(* IEC 61131-3 sources: Elmo_Master/Lasal_PRG/Welcon8Axis_EtherCAT_Test_With_RobotAxis/Class/HwControl (part 3) *)

      // safety settings
      //*********************************************************************************************
      HWC_PARA_IDX_SAFETY:

        // SubIndex
        //----------------------------------------------------------------------------------
        case SubIndex of

          //--------------------------------------------------------------------------------
          HWC_PARA_SUBIDX_SAFETY_UDP_TIME: // override cycle interval for UDP communication

            SafetyManager.GetUdpParameters(pCycleTime:=pValue$^UDINT, pTimeout:=NIL);

            Retcode := 0; // success

          //--------------------------------------------------------------------------------
          HWC_PARA_SUBIDX_SAFETY_UDP_TIMEOUT: // override timeout value for UDP communication

            SafetyManager.GetUdpParameters(pCycleTime:=NIL, pTimeout:=pValue$^UDINT);

            Retcode := 0; // success

          //--------------------------------------------------------------------------------
          else
            Retcode := -2;  // invalid SubIdx
          end_case;
    //--------------------------------------------------------------------------------
    else
      Retcode := -1;  // invalid Index
    end_case;
  end_if;

END_FUNCTION

FUNCTION GLOBAL HwControl::SetPara
	VAR_INPUT
		Index 	: DINT;
		SubIndex 	: DINT;
		Value 	: DINT;
	END_VAR
	VAR_OUTPUT
		Retcode 	: DINT;
	END_VAR

  // init returncode with invalid index
  Retcode := -1;

  // Index
  //***********************************************************************************************
  case Index of

    // safety settings
    //*********************************************************************************************
    HWC_PARA_IDX_SAFETY:

      // SubIndex
      //----------------------------------------------------------------------------------
      case SubIndex of

        //--------------------------------------------------------------------------------
        HWC_PARA_SUBIDX_SAFETY_UDP_TIME: // override cycle interval for UDP communication

          // value needs to be at least 2ms
          if Value >= 2 then
            // check if the init phase hasn't been finished yet
            if (us_InitCounter < 12) then
              SafetyManager.SetUdpParameters(pCycleTime:=(#Value)$^UDINT, pTimeout:=NIL);

              Retcode := 0; // success
            else
              Retcode := -4; // Called too late. Parameter needs to be set before the last init run.
            end_if;
          else
            Retcode := -3;  // invalid Value for this parameter
          end_if;

        //--------------------------------------------------------------------------------
        HWC_PARA_SUBIDX_SAFETY_UDP_TIMEOUT: // override timeout value for UDP communication

          // value needs to be at least 1ms
          if Value >= 1 then
            // check if the init phase hasn't been finished yet
            if (us_InitCounter < 12) then
              SafetyManager.SetUdpParameters(pCycleTime:=NIL, pTimeout:=(#Value)$^UDINT);

              Retcode := 0; // success
            else
              Retcode := -4; // Called too late. Parameter needs to be set before the last init run.
            end_if;
          else
            Retcode := -3;  // invalid Value for this parameter
          end_if;

        //--------------------------------------------------------------------------------
        else
          Retcode := -2;  // invalid SubIdx
        end_case;
  end_case;

END_FUNCTION
